TYPE ST_PLCTOROBOT_1 :
STRUCT
	arbyOutput				:ARRAY[0..31] OF BYTE;
END_STRUCT
END_TYPE

(* stored: Version 1.1.0.1, ProductVersion 3.1.4024.15
   DUT ST_PLCTOROBOT_1: Id {ee185dde-4a3f-4679-b82a-c6dc285d84b8} *)
